(* IEC 61131-3 sources: StructuredFuzzer/code_analysis/tree-sitter-structured-text, 1 file *)

(* ---- example.st ---- *)
PROGRAM My_Program
  VAR
    button1 AT %IX0.0 : BOOL := TRUE;
    button2 AT %IX0.1 : BOOL := FALSE;
    led AT %QX0.0 : BOOL;
  END_VAR
  VAR
    LED_ON : BOOL;
  END_VAR

  LED_ON := AND(button1, button2);
  IF LED_ON = TRUE THEN
    led := TRUE;
  ELSE
    led := FALSE;
  END_IF;
END_PROGRAM

CONFIGURATION STD_CONF

  RESOURCE STD_RESSOURCE ON PLC
    TASK TaskMain(INTERVAL := T#50ms,PRIORITY := 0);
    PROGRAM Inst0 WITH TaskMain : My_Program;
  END_RESOURCE
END_CONFIGURATION
